(* IEC 61131-3 sources: 2026_Projet_YGO_ExcavatriceDragage/CODE_BACKUP/CODE_20260907_ChantierWeekEnd_v0.6.43/E_CODEURS, 7 files *)

(* ---- FB_Encoder.st ---- *)
(* =======================================================================
   🔌 FB_Encoder — Objet codeur complet (1 par treuil M1/M2)
   ───────────────────────────────────────────────────────────────
   🎯 Rôle : Regrouper toute la chaine codeur derriere une interface unique :
      Abs → Homing → Scale → Safety → Reliability → Speed.
   🔌 Frontiere hardware separee HwIn/HwOut (testable).
   🔒 Homing : autorise par HomingPermit (calcule par le caller), declenche
      par HomingAtTargetM (front). La cible est fournie par le caller.
   🔒 Fiabilite : gate EncoderFault (sans Homed) calcule AVANT Speed — purge
      de vitesse au meme scan. HomedAndReliable = gate strict interlock M3.
   🧩 Defaut : Fault:ST_Fault rempli par FB_FaultCore (instFault) depuis une liste
      de causes en clair (instCauses) — pattern FB_Joystick. Ready = Enable ET pas de
      defaut late. Interlocks machine sur les faits bruts, jamais sur Fault.Latched.
   📄 Doc : DOC/AF/AF_Partie-09_Fonction_Encoder_v2.4.md
   ======================================================================= *)

FUNCTION_BLOCK PUBLIC FB_Encoder
VAR_INPUT
    // === COMMANDES & AUTORISATIONS ===
    Enable                : BOOL;        // --> [CMD] Autorisation generale FB (TRUE=Autorise)
    Reset                 : BOOL;        // --> [CMD] Acquittement defaut (front montant)

    // === AUTORISATION HOMING (calculee par le caller PRG) ===
    HomingPermit          : BOOL;        // --> [CMD] TRUE = l'operateur a le droit de homer

    // === CONSIGNES HOMING ===
    HomingAtTargetM       : BOOL;        // --> [CMD] Demande homing vers cible (front montant)
    HomingAtZero          : BOOL;        // --> [CMD] Force homing a 0.0
    ConfirmCoherence      : BOOL;        // --> [CMD] Lever le doute d'incoherence boot
    CfgHomingTargetM      : REAL;        // --> [CFG] Cible libre homing unitaire (m)
    CfgTopSensorPosM      : REAL;        // --> [CFG] Cible homing nominal capteur haut (m)
    UseDynamicTarget      : BOOL;        // --> [CMD] Active cible dynamique
    DynamicHomingTargetM  : REAL;       // --> [CFG] Cible dynamique de referencement (m)

    // === CAPTEURS PHYSIQUES ===
    TopPositionSensor     : BOOL;        // --> [HW]  Capteur physique position haute unique

    // === BUS ETHERCAT & CAPTEUR HW (frontiere testable) ===
    HwIn                  : ST_fbEncoder_HwIn; // --> [HW] Retours hardware codeur

    // === MECANIQUE (constantes) ===
    PointsPerRev          : UDINT := 8192; // --> [CFG] Resolution codeur (pts/tour)
    CableM_PerRev         : REAL := 2.0;   // --> [CFG] Developpement cable par tour (m/tour)

    // === REGLAGES & CONFIGURATION ===
    Cfg                   : ST_fbEncoder_Cfg; // --> [CFG] Mode de confirmation preset
    PositionMinM          : REAL := -99.0; // --> [CFG] Plafond bornage physique bas (m)
    PositionMaxM          : REAL := 99.0;  // --> [CFG] Plafond bornage physique haut (m)
    BypassGlobal          : BOOL := FALSE; // --> [TST] Neutralisation defauts pour mise en service
END_VAR
VAR_OUTPUT
    // === ETATS IEC & SYNOPTIQUE ===
    Ready                 : BOOL;        // <-- [STAT] FB pret a fonctionner (Enable ET pas de defaut late)
    Fault                 : ST_Fault;    // <-- [DIAG] Brique defaut socle (live + latchee), remplie par FB_FaultCore

    // === FRONTIERE HW SORTIE (testable) ===
    HwOut                 : ST_fbEncoder_HwOut; // <-- [ACT] Ordres hardware codeur (preset)

    // === MESURES CONDITIONNEES (struct frontiere) ===
    Measurement           : ST_fbEncoder_Measurement; // <-- [BUS] Mesures + statuts (interface)

    // === ETATS CODEUR ===
    Homed                 : BOOL;        // <-- [STAT] Codeur reference (sortie homing)
    HomingSuspect         : BOOL;        // <-- [DIAG] Incoherence redemarrage a lever
    EncoderFault          : BOOL;        // <-- [SAFE] Gate general fiabilite (sans Homed)
    HomedAndReliable      : BOOL;        // <-- [STAT] Gate strict M3 : dispo ET ref ET pas incoherent
    PresetConfirmationFailed : BOOL;     // <-- [DIAG] Latch derniere verification preset echouee
END_VAR
VAR
    // === SOUS-INSTANCES FB (chaine codeur complete) ===
    instAbs        : FB_Encoder_Abs;          // * [INST] Acquisition brute codeur EtherCAT
    instHoming     : FB_Encoder_Homing;       // * [INST] Referencement (homing) nominal/unitaire
    instScale      : FB_Encoder_Scale;        // * [INST] Mise a l'echelle points -> metres
    instSafety     : FB_Encoder_Safety;       // * [INST] Bornage & coherence mesure
    instRel        : FB_EncoderReliability;   // * [INST] Gates de fiabilite
    instSpeed      : FB_Encoder_SpeedMeasure; // * [INST] Calcul vitesse cable
    instFault      : FB_FaultCore;            // * [INST] Socle de defaut (liste de causes -> ST_Fault)
    instCauses     : ARRAY[0..15] OF ST_FaultCause; // . [LOC] Liste des causes pour le socle FB_FaultCore
END_VAR
VAR_IN_OUT
    // === CALIBRATION PERSISTANTE (externe RETAIN, jamais membre) ===
    Calib                  : ST_Encoder_Calib; // <-> [BUS] Calibration RETAIN du treuil
END_VAR

{region "§1 Gate neutralisation"}
IF NOT Enable THEN
    Ready := FALSE;
    Measurement.RawPos := 0; Measurement.EncoderAvailable := FALSE;
    Measurement.CablePosM := 0.0; Measurement.CablePosMSafe := 0.0; Measurement.EncoderIncoherent := FALSE;
    Measurement.Speed_Mps := 0.0; Measurement.SignedSpeed_Mps := 0.0; Measurement.SpeedValid := FALSE;
    Measurement.HomingFault.Error := FALSE; Measurement.HomingFault.ErrorId := 0;
    Measurement.HomingLifecycle.Busy := FALSE; Measurement.HomingLifecycle.Done := FALSE;
    Measurement.AbsFault.Error := FALSE;    Measurement.AbsFault.ErrorId := 0;
    EncoderFault := TRUE;
    HomedAndReliable := FALSE;
    // Frontiere HW sortie : aucun ordre preset publie hors autorisation
    // (sinon PRG_02_Acquisition relaie une valeur perimee au codeur absolu -> preset parasite, reference corrompue)
    HwOut.PresetTriggerCmd := 0; HwOut.CodeSeqTriggerCmd := 0; HwOut.PresetValueOut := 0;
    // Reference connue MAINTENUE depuis Calib (RETAIN) meme FB desactive (AF09 §4) :
    // un FB desactive ne doit pas faire perdre la reference aux consommateurs aval (PRG_04, FB_Encoder_Scale).
    Homed := Calib.Homed;
    HomingSuspect := Calib.HomingSuspect;
    Measurement.HomingRefRaw := Calib.HomingRefRaw;
    // PresetConfirmationFailed est un diagnostic latch : il reste gele hors Enable
    // et ne doit pas etre efface par ce gate (AC3).
    // Socle appele meme Enable=FALSE : maintient le latch non acquitte et traite le Reset
    // hors autorisation (AC4). Les causes ne sont pas evaluees (Enable=FALSE -> vue live a 0),
    // les latches sont preserves.
    instFault(Enable := FALSE, Reset := Reset, Causes := instCauses);
    Fault := instFault.Fault;
    RETURN;
END_IF;
Ready := TRUE;
{endregion}

{region "§2 Abs"}
    instAbs(
    Enable              := Enable,
    Reset               := Reset,
    RawPosIn            := HwIn.RawPosIn,
    AlarmsIn            := HwIn.AlarmsIn,
    WarningsIn          := HwIn.WarningsIn,
    SlaveOperational    := HwIn.SlaveOperational,
    PresetRequest       := instHoming.PresetRequest,
    PresetValue         := instHoming.PresetValue,
    PointsPerRev        := PointsPerRev
);
{endregion}

{region "§3 Homing"}
instHoming(
    Enable               := Enable,
    Reset                := Reset,
    Home                 := HomingAtTargetM,
    HomingPermit         := HomingPermit,
    BtnConfirmCoherence  := ConfirmCoherence,
    UseDynamicTarget     := UseDynamicTarget,
    DynamicHomingTargetM := DynamicHomingTargetM,
    CfgHomingTargetM     := CfgHomingTargetM,
    CfgTopSensorPosM     := SEL(HomingAtZero, CfgTopSensorPosM, 0.0),
    TopPositionSensor    := TopPositionSensor,
    RawPos               := instAbs.RawPos,
    EncoderAvailable     := instAbs.EncoderAvailable,
    PresetStatusBit      := HwIn.PresetStatusBit,
    Cfg                  := Cfg,
    PointsPerRev         := PointsPerRev,
    MultiTurnRevsMax     := 4096,
    CableM_PerRev        := CableM_PerRev,
    BypassGlobal         := BypassGlobal,
    Calib                := Calib
);
{endregion}

{region "§4 Scale"}
instScale(
    RawPos       := instAbs.RawPos,
    HomingRefRaw := instHoming.HomingRefRaw,
    CableM_PerRev := CableM_PerRev,
    PointsPerRev := PointsPerRev
);
{endregion}

{region "§5 Safety"}
instSafety(
    Enable             := Enable,
    Reset              := Reset,
    CablePosM          := instScale.CablePosM,
    HomingSuspect      := instHoming.HomingSuspect,
    PositionMinM       := PositionMinM,
    PositionMaxM       := PositionMaxM,
    BypassGlobal       := BypassGlobal
);
{endregion}

{region "§6 Reliability"}
instRel(
    EncoderAvailable  := instAbs.EncoderAvailable,
    Homed             := instHoming.Homed,
    EncoderIncoherent := instSafety.EncoderIncoherent
);
{endregion}

{region "§7 Speed"}
instSpeed(
    Enable        := Enable,
    Reset         := Reset,
    SpdValueIn    := HwIn.SpdValueIn,
    PositionValid := NOT instRel.EncoderFault,
    CableM_PerRev := CableM_PerRev
);
{endregion}

{region "§8 Remplissage struct et synthese"}
Measurement.RawPos            := instAbs.RawPos;
Measurement.EncoderAvailable  := instAbs.EncoderAvailable;
Measurement.CablePosM         := instSafety.CablePosMSafe;
Measurement.CablePosMSafe     := instSafety.CablePosMSafe;
Measurement.EncoderIncoherent := instSafety.EncoderIncoherent;
Measurement.Speed_Mps         := instSpeed.Speed_Mps;
Measurement.SignedSpeed_Mps   := instSpeed.SignedSpeed_Mps;
Measurement.SpeedValid        := instSpeed.Valid;
Measurement.HomingFault        := instHoming.Fault;
Measurement.HomingLifecycle    := instHoming.Lifecycle;
Measurement.AbsFault           := instAbs.Fault;
Measurement.HomingRefRaw      := instHoming.HomingRefRaw;

// Frontiere HW sortie (preset)
HwOut.PresetTriggerCmd := instAbs.PresetTriggerCmd;
HwOut.CodeSeqTriggerCmd := instAbs.CodeSeqTriggerCmd;
HwOut.PresetValueOut    := instAbs.PresetValueOut;

// Etats codeur
Homed            := instHoming.Homed;
HomingSuspect    := instHoming.HomingSuspect;
EncoderFault     := instRel.EncoderFault;
HomedAndReliable := instRel.HomedAndReliable;
PresetConfirmationFailed := instHoming.PresetConfirmationFailed;

// Synthese statut facade : brique defaut socle (Fault:ST_Fault), pattern FB_Joystick.
// Causes exprimees en CLAIR (ST_FaultCause), alimentees UNIQUEMENT depuis les sorties
// publiques des sous-FB (encapsulation stricte, jamais de lecture VAR interne).
//   - Cause 0/1 : LIVE (Latching=FALSE) -> Fault.Error, retombe seule.
//   - Cause 2   : LATCHED (Latching=TRUE) -> arme Fault.Latched, acquittee au Reset front.
// Interlock machine toujours sur les faits bruts (EncoderFault, HomedAndReliable,
// EncoderIncoherent), jamais sur Fault.Latched (conservation).
instCauses[0].Active := NOT instAbs.EncoderAvailable; instCauses[0].Latching := FALSE;
instCauses[0].Texte := 'Perte materiel / communication codeur EtherCAT';
instCauses[1].Active := instSafety.EncoderIncoherent; instCauses[1].Latching := FALSE;
instCauses[1].Texte := 'Incoherence mesure / saut de position codeur';
instCauses[2].Active := instHoming.PresetConfirmationFailed; instCauses[2].Latching := TRUE;
instCauses[2].Texte := 'Echec confirmation transaction preset codeur';

// Socle appele APRES le pipeline : causes du scan courant, aucun scan de retard (AC4).
instFault(Enable := Enable, Reset := Reset, Causes := instCauses);
Fault := instFault.Fault;     // source de verite = socle
Ready := Enable AND NOT Fault.Latched;
{endregion}

(* ---- FB_Encoder_Abs.st ---- *)
(* =======================================================================
   🔌 FB_Encoder_Abs — Acquisition codeur absolu (accès bus EtherCAT)
   ───────────────────────────────────────────────────────────────
   🎯 Rôle : Accès bus EtherCAT, extraction positions brutes et séquence de Preset SDO
   🔒 Polarité : EncoderAvailable=TRUE si communication bus et esclave OK
   🔌 Architecture : Module d'acquisition codeur absolu
   📄 Doc métier : DOC/AF/AF_Partie-09_Fonction_Encoder_v2.4.md
   ======================================================================= *)

// === DECLARATION (à coller dans la partie déclaration du POU FB_Encoder_Abs) ===

FUNCTION_BLOCK PUBLIC FB_Encoder_Abs
VAR_INPUT
    // === COMMANDES & AUTORISATIONS ===
    Enable              : BOOL;        // --> [CMD] Autorisation generale FB (TRUE=Autorise)
    Reset               : BOOL;        // --> [CMD] Acquittement defaut (front montant)
    PresetRequest       : BOOL;        // --> [CMD] Demande de preset (front montant)

    // === BUS ETHERCAT & CAPTEUR HW ===
    RawPosIn            : UDINT;       // --> [HW]  Position brute EtherCAT
    AlarmsIn            : UINT;        // --> [HW]  Codes alarmes bruts EtherCAT
    WarningsIn          : UINT;        // --> [HW]  Codes avertissements bruts EtherCAT
    SlaveOperational    : BOOL;        // --> [HW]  Statut esclave EtherCAT operationnel

    // === PARAMETRES & REGLAGES ===
    PointsPerRev        : UDINT := 8192; // --> [CFG] Resolution codeur (pts/tour)
    PresetValue         : UDINT;       // --> [CFG] Valeur cible de preset
    PresetTimeout       : TIME := T#2s;// --> [CFG] Temporisation max attente preset
    PresetTolerancePts  : UDINT := 10; // --> [CFG] Tolerance relecture post-preset (pts)
END_VAR
VAR_OUTPUT
    // === ETATS IEC & SYNOPTIQUE ===
    Ready               : BOOL;        // <-- [STAT] FB pret a fonctionner
    // 🧩 Statut transverse (forme cible ST_Fault)
    Fault               : ST_Fault;

    // === MESURES & DONNEES CODEUR ===
    RawPos              : UDINT;       // <-- [DIAG] Position brute gelee si non disponible
    EncoderAvailable    : BOOL;        // <-- [STAT] Codeur operationnel et disponible
    AngleRaw            : UINT;        // <-- [DIAG] Angle brut sur un tour (MOD PointsPerRev)
    TurnCount           : UDINT;       // <-- [DIAG] Nombre de tours bruts (RawPos / PointsPerRev)

    // === COMMANDES & ECHANGE BUS ETHERCAT ===
    PresetTriggerCmd    : WORD;        // <-- [ACT]  Ordre declenchement preset vers PDO Rx
    CodeSeqTriggerCmd   : WORD;        // <-- [ACT]  Ordre sequence code vers PDO Rx
    PresetValueOut      : UDINT;       // <-- [ACT]  Valeur de preset transmise au PDO Rx
END_VAR
VAR
    // === DETECTEURS DE FRONT ===
    ResetEdge           : R_TRIG;      // . [LOC] Detecteur front montant Reset
    PresetReqEdge       : R_TRIG;      // . [LOC] Detecteur front montant PresetRequest

    // === TEMPORISATEURS INTERNES ===
    PresetTimer         : TON;         // . [LOC] Temporisateur timeout sequence preset
    PresetTimerVisual   : TON;         // . [LOC] Temporisateur maintien visuel impulsion (500ms)

    // === VARIABLES INTERNES DE CALCUL & ETAT ===
    PresetSeqStep       : INT;         // . [LOC] Etape sequence preset (0:IDLE, 1:PULSE/WAIT)
    RawDiff             : DINT;        // . [LOC] Ecart signe entre RawPos et PresetValueOut
    PresetCompleted     : BOOL;        // . [LOC] Fait de fin de maintien preset (un scan)
    PresetTimeoutError  : BOOL;        // . [LOC] Latch interne timeout séquence preset

    // === SOCLE DEFAUT (FB_FaultCore) ===
    instFault           : FB_FaultCore;                   // * [INST] Socle défaut transverse
    instCauses          : ARRAY[0..15] OF ST_FaultCause;  // . [LOC] Table des causes nommées
END_VAR

// === IMPLEMENTATION (à coller dans le corps ST du POU FB_Encoder_Abs) ===

{region "§1 Causes & Socle Défaut (évalué en continu)"}
// 🔑 1. RESET FRONT
ResetEdge(CLK := Reset);

// 🔍 2. DIAGNOSTIC BUS / ALARME (Cause 0 : live)
instCauses[0].Active   := (AlarmsIn <> 0) OR NOT SlaveOperational;
instCauses[0].Latching := FALSE;
instCauses[0].Texte    := 'Defaut communication EtherCAT codeur absolu';

// ⏱️ 3. TIMEOUT PRESET (Cause 1 : latched)
IF ResetEdge.Q AND (PresetSeqStep = 0) THEN
    PresetTimeoutError := FALSE;
END_IF;
instCauses[1].Active   := PresetTimeoutError;
instCauses[1].Latching := TRUE;
instCauses[1].Texte    := 'Timeout sequence preset SDO codeur';

// Appel du socle de défaut
instFault(Enable := Enable, Reset := Reset, Causes := instCauses);
Fault := instFault.Fault;

EncoderAvailable := NOT instCauses[0].Active;
{endregion}

{region "§2 Gate neutralisation"}
// 🛑 2. GATE
IF NOT Enable THEN
    EncoderAvailable := FALSE;
    Ready := FALSE;
    PresetTriggerCmd := 0; CodeSeqTriggerCmd := 0; PresetValueOut := 0;
    PresetSeqStep := 0;
    PresetCompleted := FALSE;
    PresetTimer(IN := FALSE, PT := PresetTimeout);
    PresetTimerVisual(IN := FALSE, PT := T#500MS);
    // RawPos, AngleRaw et TurnCount sont volontairement gelés hors Enable
    // (AF09 F09.01 / AC5) : aucune lecture bus ni remise a zero dans ce gate.
    RETURN;
END_IF;

Ready := Enable AND NOT Fault.Latched;
{endregion}

{region "§3 Lecture position"}
// 📥 3. LECTURE POSITION — GELER SUR DOUTE (Partie10 §6)
// Si EncoderAvailable=FALSE : RawPos/AngleRaw/TurnCount conservent leur dernière valeur (pas de RETURN
// global ici pour ne pas geler aussi la séquence preset/l'état — seule la lecture est gelée).
IF EncoderAvailable THEN
    RawPos := RawPosIn;   // Sens de comptage géré côté codeur (CoE 6000h bit0, startup parameter CODESYS) — voir Partie10 §3bis. Plus de calcul ici.
    AngleRaw := UDINT_TO_UINT(RawPos MOD PointsPerRev);
    TurnCount := RawPos / PointsPerRev;
END_IF;
{endregion}

{region "§4 Séquence preset"}
// 🔧 4. SÉQUENCE PRESET (écriture bus)
// PresetTriggerCmd := 2 déclenche le référencement à PresetValue (valeur de commande, pas un
// masque de bits). CodeSeqTriggerCmd : rôle non identifié — laissé à 0, PAS piloté tant que sa
// fonction n'est pas confirmée. Ne jamais lui donner une valeur arbitraire.
PresetReqEdge(CLK := PresetRequest);
PresetCompleted := FALSE;
CodeSeqTriggerCmd := 0;                 // non piloté — rôle inconnu, voir note ci-dessus
CASE PresetSeqStep OF
    0: // IDLE
        PresetTriggerCmd := 0;
        IF PresetReqEdge.Q AND EncoderAvailable THEN
            PresetValueOut := PresetValue;
            PresetSeqStep := 1;
            PresetTimer(IN := TRUE, PT := PresetTimeout);
        END_IF;
    1: // Déclenchement preset (laissé actif pendant 0.5s pour confort visuel en simulation/bus)
        PresetTriggerCmd := 2;   // Référence le codeur à PresetValueOut
        RawDiff := UDINT_TO_DINT(RawPos) - UDINT_TO_DINT(PresetValueOut);
        IF ABS(RawDiff) <= UDINT_TO_DINT(PresetTolerancePts) THEN
            PresetTimer(IN := FALSE, PT := PresetTimeout);
            PresetTimerVisual(IN := TRUE, PT := T#500MS);
            IF PresetTimerVisual.Q THEN
                PresetTriggerCmd := 0;
                PresetCompleted := TRUE;
                PresetSeqStep := 0;
                PresetTimerVisual(IN := FALSE, PT := T#500MS);
            END_IF;
        ELSIF PresetTimer.Q THEN
            PresetTriggerCmd := 0;
            PresetTimeoutError := TRUE;
            PresetSeqStep := 0;
            PresetTimer(IN := FALSE, PT := PresetTimeout);
            PresetTimerVisual(IN := FALSE, PT := T#500MS);
        END_IF;
END_CASE;
{endregion}

(* ---- FB_Encoder_Homing.st ---- *)
(* =======================================================================
   ⚙️ FB_Encoder_Homing — Référencement codeur nominal ou unitaire
   ───────────────────────────────────────────────────────────────
   🎯 Rôle : Séquence de référencement nominal (capteur haut) ou unitaire (MAINT_N2)
   🔒 Polarité : Homed=TRUE dès qu'un référencement valide est enregistré
   🔌 Architecture : Expose ST_Encoder_Calib en VAR_IN_OUT
   📄 Doc métier : DOC/AF/AF_Partie-09_Fonction_Encoder_v2.4.md
   ======================================================================= *)

// === DECLARATION (à coller dans la partie déclaration du POU FB_Encoder_Homing) ===

FUNCTION_BLOCK PUBLIC FB_Encoder_Homing
VAR_INPUT
    // === COMMANDES & AUTORISATIONS ===
    Enable                 : BOOL;        // --> [CMD] Autorisation generale FB (TRUE=Autorise)
    Reset                  : BOOL;        // --> [CMD] Acquittement defaut (front montant)
    Home                   : BOOL;        // --> [CMD] Demande de referencement (front)
    HomingPermit           : BOOL;        // --> [CMD] Autorisation de homer (calculee par le caller)
    BtnConfirmCoherence    : BOOL;        // --> [CMD] Levee de doute d'incoherence au boot (front)

    // === CIBLES & CONFIGURATION HOMING ===
    CfgHomingTargetM       : REAL;        // --> [CFG] Cible libre homing unitaire (m)
    UseDynamicTarget       : BOOL := FALSE; // --> [CFG] Activation cible dynamique
    DynamicHomingTargetM   : REAL := 0.0; // --> [CFG] Cible dynamique de referencement (m)
    CfgTopSensorPosM       : REAL := 8.5; // --> [CFG] Cible homing nominal capteur haut (m)

    // === RETOURS HW & CAPTEURS ===
    TopPositionSensor      : BOOL;        // --> [HW]  Capteur physique position haute unique
    // === MESURES & RETOURS FB CODEUR ABSOLU ===
    RawPos                 : UDINT;       // --> [HW]  Position brute codeur (sortie FB_Encoder_Abs)
    EncoderAvailable       : BOOL;        // --> [HW]  Codeur absolu disponible et valide
    PresetStatusBit        : BOOL;        // --> [HW]  Bit d'etat preset optionnel, FALSE si non cable

    // === REGLAGES TRANSACTION PRESET ===
    Cfg                    : ST_fbEncoder_Cfg; // --> [CFG] Mode de confirmation preset

    // === CARACTERISTIQUES MECANIQUES & BUS ===
    PointsPerRev           : UDINT := 8192; // --> [CFG] Resolution codeur (pts/tour)
    MultiTurnRevsMax       : UDINT := 4096; // --> [CFG] Capacite multitour max codeur (tours)
    CableM_PerRev          : REAL := 2.0;   // --> [CFG] Perimetre tambour / developpement cable (m/tour)

    // === TESTS & BYPASS ===
    BypassGlobal           : BOOL := FALSE; // --> [TST] Neutralisation securites pour mise en service
END_VAR
VAR_OUTPUT
    // === ETATS IEC & SYNOPTIQUE ===
    Ready                  : BOOL;        // <-- [STAT] FB pret a fonctionner
    // 🧩 Statut transverse (forme cible ST_Fault)
    Fault                  : ST_Fault;
    // 🧩 Cycle de vie (forme cible ST_Lifecycle)
    Lifecycle              : ST_Lifecycle;

    // === COMMANDES VERS FB_ENCODER_ABS ===
    PresetRequest          : BOOL;        // <-- [ACT]  Pulse demande d'ecriture preset SDO
    PresetValue            : UDINT;       // <-- [ACT]  Valeur de cible brute pour preset SDO

    // === RESULTATS & MEMOIRE CALIBRATION ===
    Homed                  : BOOL;        // <-- [STAT] Codeur pagine et referencie
    HomingSuspect          : BOOL;        // <-- [DIAG] Incoherence redemarrage a lever
    HomingRefRaw           : UDINT;       // <-- [DIAG] Offset de reference brut calcule
    PresetConfirmationFailed : BOOL;      // <-- [DIAG] Latch derniere verification preset echouee
END_VAR
VAR_IN_OUT
    // === STRUCTURE DE CALIBRATION PERSISTANTE ===
    Calib                  : ST_Encoder_Calib; // <-> [BUS] Structure de calibration RETAIN
END_VAR
VAR
    // === DETECTEURS DE FRONT ===
    ResetEdge              : R_TRIG;      // . [LOC] Detecteur front montant Reset
    HomeEdge               : R_TRIG;      // . [LOC] Detecteur front montant Home
    ConfirmCoherenceEdge   : R_TRIG;      // . [LOC] Detecteur front montant BtnConfirmCoherence
    TopSensorEdge          : R_TRIG;      // . [LOC] Detecteur front montant TopPositionSensor
    DynamicTargetEdge      : R_TRIG;      // . [LOC] Detecteur front montant UseDynamicTarget

    // === ETATS & DRAPEAUX INTERNES ===
    InitDone               : BOOL;        // . [LOC] Controle incoherence boot effectue
    HomingModeOk           : BOOL;        // . [LOC] Mode de fonctionnement valide pour homing
    NominalHomingTrigger   : BOOL;        // . [LOC] Condition de declenchement homing nominal
    UnitaryHomingTrigger   : BOOL;        // . [LOC] Condition de declenchement homing unitaire
    DynamicHomingTrigger   : BOOL;        // . [LOC] Condition de declenchement homing dynamique
    HomingTrigger          : BOOL;        // . [LOC] Synthese declenchement homing
    PresetVerificationActive : BOOL;      // . [LOC] Verification preset en attente
    PresetConfirmed        : BOOL;        // . [LOC] Resultat du mode de confirmation selectionne

    // === DRAPEAUX DEFAUTS INTERNES ===
    HomingModeError        : BOOL;        // . [LOC] Latch erreur mode
    TargetOutOfRangeError  : BOOL;        // . [LOC] Latch cible hors limites
    PresetFailError        : BOOL;        // . [LOC] Latch échec preset
    BootIncoherentError    : BOOL;        // . [LOC] Latch incohérence boot

    // === VARIABLES DE CALCUL ===
    TargetPoints           : DINT;        // . [LOC] Ecart cible converti en points
    TargetPositionM        : REAL;        // . [LOC] Cible retenue en metres
    RawDiffRestart         : DINT;        // . [LOC] Ecart brut de position au redemarrage
    PendingHomingRefRaw    : UDINT;       // . [LOC] Reference candidate, non publiee avant succes
    CandidateRawDiff       : DINT;        // . [LOC] Ecart brut de la mesure candidate
    CandidateCablePosM     : REAL;        // . [LOC] Position candidate calculee avant commit
    ReadbackOk             : BOOL;        // . [LOC] Mesure candidate dans la tolerance
    StatusBitOk            : BOOL;        // . [LOC] Etat du bit optionnel de confirmation
    PresetVerifyTimer      : TON;         // . [LOC] Temporisation historique de verification 500ms

    // === SOCLE DEFAUT (FB_FaultCore) ===
    instFault              : FB_FaultCore;                   // * [INST] Socle défaut transverse
    instCauses             : ARRAY[0..15] OF ST_FaultCause;  // . [LOC] Table des causes nommées
END_VAR

VAR CONSTANT
    // === TOLERANCE & TEMPORISATION TRANSACTION ===
    CST_HomingVerifyToleranceM : REAL := 0.010; // Tolerance mesure cible (m)
    CST_PresetVerifyTime        : TIME := T#50MS; // Latence historique avant relecture
END_VAR

// === IMPLEMENTATION (à coller dans le corps ST du POU FB_Encoder_Homing) ===

{region "§1 Causes & Socle Défaut (évalué en continu)"}
// 🔑 1. FRONTS
ResetEdge(CLK := Reset);
HomeEdge(CLK := Home);
ConfirmCoherenceEdge(CLK := BtnConfirmCoherence);

// Effacement des latches d'erreur sur Reset conscient
IF ResetEdge.Q THEN
    PresetConfirmationFailed := FALSE;
    HomingModeError := FALSE;
    TargetOutOfRangeError := FALSE;
    PresetFailError := FALSE;
END_IF;

// Levée de doute incohérence boot (BtnConfirmCoherence)
IF ConfirmCoherenceEdge.Q AND HomingPermit THEN
    Calib.HomingSuspect := FALSE;
    BootIncoherentError := FALSE;
END_IF;

// Configuration des causes nommées
instCauses[0].Active   := HomingModeError;
instCauses[0].Latching := TRUE;
instCauses[0].Texte    := 'Homing non autorise dans ce mode';

instCauses[1].Active   := TargetOutOfRangeError;
instCauses[1].Latching := TRUE;
instCauses[1].Texte    := 'Cible de homing hors plage';

instCauses[2].Active   := PresetFailError;
instCauses[2].Latching := TRUE;
instCauses[2].Texte    := 'Echec confirmation transaction preset';

instCauses[3].Active   := BootIncoherentError;
instCauses[3].Latching := TRUE;
instCauses[3].Texte    := 'Incoherence position codeur au demarrage';

// Appel du socle de défaut
instFault(Enable := Enable, Reset := Reset, Causes := instCauses);
Fault := instFault.Fault;
{endregion}

{region "§2 Gate neutralisation"}
// 🛑 2. GATE — neutralisation ; on continue toutefois d'exposer le dernier état RETAIN connu
// (FB_Encoder_Scale a besoin de HomingRefRaw même si ce FB est désactivé)
IF NOT Enable THEN
    PresetRequest := FALSE;
    PresetValue := 0;
    Ready := FALSE;
    Lifecycle.Busy := FALSE;
    Lifecycle.Done := FALSE;
    InitDone := FALSE;   // Force un nouveau contrôle à la prochaine activation
    PresetVerificationActive := FALSE;
    PresetVerifyTimer(IN := FALSE, PT := CST_PresetVerifyTime);
    Homed := Calib.Homed;
    HomingSuspect := Calib.HomingSuspect;
    HomingRefRaw := Calib.HomingRefRaw;
    // PresetConfirmationFailed est un diagnostic latch : il est gelé hors Enable
    RETURN;
END_IF;

Ready := Enable AND NOT Fault.Latched;
{endregion}

{region "§3 Cohérence au redémarrage"}
// 🔍 3. COHÉRENCE AU REDÉMARRAGE — une fois par session Enable, dès que le codeur répond
IF NOT InitDone THEN
    IF EncoderAvailable THEN
        RawDiffRestart := UDINT_TO_DINT(RawPos) - UDINT_TO_DINT(Calib.LastKnownRawPos);
        IF Calib.Homed AND (ABS(RawDiffRestart) > UDINT_TO_DINT(Calib.RestartCoherenceTolerancePts)) THEN
            Calib.HomingSuspect := TRUE;
            BootIncoherentError := TRUE;
        END_IF;
        InitDone := TRUE;
    END_IF;
END_IF;
{endregion}

{region "§4 Demande et déclenchement homing"}
// ⚙️ 4. DEMANDE & DÉCLENCHEMENT HOMING
PresetRequest := FALSE;
PresetValue := 0;
TopSensorEdge(CLK := TopPositionSensor);
DynamicTargetEdge(CLK := UseDynamicTarget);

HomingModeOk := HomingPermit;

IF HomeEdge.Q AND NOT HomingModeOk THEN
    HomingModeError := TRUE;
END_IF;

NominalHomingTrigger := HomingModeOk AND NOT UseDynamicTarget
                         AND ((Home AND TopSensorEdge.Q) OR (HomeEdge.Q AND TopPositionSensor));

UnitaryHomingTrigger := HomingModeOk AND NOT UseDynamicTarget AND HomeEdge.Q;

DynamicHomingTrigger := HomingModeOk AND (DynamicTargetEdge.Q OR (UseDynamicTarget AND HomeEdge.Q));

HomingTrigger := (NominalHomingTrigger OR UnitaryHomingTrigger OR DynamicHomingTrigger)
                 AND NOT PresetVerificationActive;

IF HomingTrigger THEN
    IF UseDynamicTarget THEN
        TargetPositionM := DynamicHomingTargetM;
    ELSIF NominalHomingTrigger THEN
        TargetPositionM := CfgTopSensorPosM;
    ELSE
        TargetPositionM := CfgHomingTargetM;
    END_IF;

    // Bornage obligatoire avant écriture (CODE_QUALITY_STANDARDS §6) [-99;+99] m
    IF (TargetPositionM < -99.0) OR (TargetPositionM > 99.0) THEN
        TargetOutOfRangeError := TRUE;
    ELSE
        TargetPoints := REAL_TO_DINT(TargetPositionM * UDINT_TO_REAL(PointsPerRev) / CableM_PerRev);
        PendingHomingRefRaw := DINT_TO_UDINT(UDINT_TO_DINT(RawPos) - TargetPoints);
        PresetValue := RawPos;
        PresetRequest := TRUE;
        PresetVerificationActive := TRUE;
        Lifecycle.Done := FALSE;
    END_IF;
END_IF;
{endregion}

{region "§5 Suivi de transaction preset"}
// ⏳ 5. SUIVI DE LA TRANSACTION PRESET
PresetVerifyTimer(IN := PresetVerificationActive, PT := CST_PresetVerifyTime);
IF PresetVerificationActive AND PresetVerifyTimer.Q THEN
    CandidateRawDiff := UDINT_TO_DINT(RawPos) - UDINT_TO_DINT(PendingHomingRefRaw);
    IF PointsPerRev <> 0 THEN
        CandidateCablePosM := DINT_TO_REAL(CandidateRawDiff) * CableM_PerRev / UDINT_TO_REAL(PointsPerRev);
    ELSE
        CandidateCablePosM := 0.0;
    END_IF;
    ReadbackOk := ABS(CandidateCablePosM - TargetPositionM) <= CST_HomingVerifyToleranceM;
    StatusBitOk := PresetStatusBit;

    CASE Cfg.PresetConfirmMode OF
        E_PresetConfirmMode.READBACK_ONLY:
            PresetConfirmed := ReadbackOk;
        E_PresetConfirmMode.READBACK_AND_STATUSBIT:
            PresetConfirmed := ReadbackOk AND StatusBitOk;
        E_PresetConfirmMode.STATUSBIT_ONLY:
            PresetConfirmed := StatusBitOk;
        ELSE
            PresetConfirmed := FALSE;
    END_CASE;

    IF PresetConfirmed THEN
        Calib.HomingRefRaw := PendingHomingRefRaw;
        Calib.Homed := TRUE;
        Calib.HomingSuspect := FALSE;
        Calib.LastKnownRawPos := RawPos;
        PresetConfirmationFailed := FALSE;
        PresetFailError := FALSE;
        Lifecycle.Done := TRUE;
    ELSE
        Calib.HomingSuspect := TRUE;
        PresetConfirmationFailed := TRUE;
        PresetFailError := TRUE;
        Lifecycle.Done := FALSE;
    END_IF;

    PresetVerificationActive := FALSE;
    PresetVerifyTimer(IN := FALSE, PT := CST_PresetVerifyTime);
END_IF;
{endregion}

{region "§6 Sorties état & calibration"}
// 📤 6. SORTIES ÉTAT & CALIBRATION
IF EncoderAvailable AND NOT PresetVerificationActive THEN
    Calib.LastKnownRawPos := RawPos;
END_IF;

Lifecycle.Busy := PresetVerificationActive;
Homed := Calib.Homed AND NOT Calib.HomingSuspect;
HomingSuspect := Calib.HomingSuspect;
HomingRefRaw := Calib.HomingRefRaw;
{endregion}

(* ---- FB_Encoder_Safety.st ---- *)
(* =======================================================================
   🛡️ FB_Encoder_Safety — Bornage physique & surveillance cohérence
   ───────────────────────────────────────────────────────────────
   🎯 Rôle : Bornage physique absolu [-99; +99]m et relais d'incohérence redémarrage
   🔒 Polarité : EncoderIncoherent=TRUE en cas de hors bornes ou HomingSuspect
   🛡️ Sécurité : Verrouillage de la position câble sûre
   📄 Doc métier : DOC/AF/AF_Partie-09_Fonction_Encoder_v2.4.md
   ======================================================================= *)

FUNCTION_BLOCK PUBLIC FB_Encoder_Safety
VAR_INPUT
    // === COMMANDES & AUTORISATIONS ===
    Enable                : BOOL;        // --> [CMD] Autorisation generale FB (TRUE=Autorise)
    Reset                 : BOOL;        // --> [CMD] Acquittement defaut (front montant)

    // === MESURES & ALERTE HOMING ===
    CablePosM             : REAL;        // --> [HW]  Position calculee (m, sortie FB_Encoder_Scale)
    HomingSuspect         : BOOL;        // --> [SAFE] Alerte incoherence redemarrage (FB_Encoder_Homing)

    // === REGLAGES & BORNES PHYSIQUES ===
    PositionMinM          : REAL := -99.0; // --> [CFG] Plafond bornage physique bas (m)
    PositionMaxM          : REAL := 99.0;  // --> [CFG] Plafond bornage physique haut (m)

    // === TESTS & BYPASS ===
    BypassGlobal          : BOOL := FALSE; // --> [TST] Neutralisation defaut de bornage pour mise en service
END_VAR
VAR_OUTPUT
    // === ETATS IEC & SYNOPTIQUE ===
    Ready                 : BOOL;        // <-- [STAT] FB pret a fonctionner
    // 🧩 Statut transverse (forme cible ST_Fault)
    Fault                 : ST_Fault;

    // === MESURES SURE & SECURITE ===
    CablePosMSafe         : REAL;        // <-- [DIAG] Position cable instantanee transmise (m)
    EncoderIncoherent     : BOOL;        // <-- [SAFE] Incoherence ou hors bornes (TRUE = defaut)
END_VAR
VAR
    // === DETECTEURS DE FRONT ===
    ResetEdge             : R_TRIG;      // . [LOC] Detecteur front montant Reset

    // === SOCLE DEFAUT (FB_FaultCore) ===
    instFault             : FB_FaultCore;                   // * [INST] Socle défaut transverse
    instCauses            : ARRAY[0..15] OF ST_FaultCause;  // . [LOC] Table des causes nommées
END_VAR

// === IMPLEMENTATION ===

{region "§1 Causes & Socle Défaut (évalué en continu)"}
// 🔑 1. RESET FRONT
ResetEdge(CLK := Reset);

// 🔍 2. SURVEILLANCE BORNAGE & INCOHÉRENCE BOOT
instCauses[0].Active   := NOT BypassGlobal AND ((CablePosM < PositionMinM) OR (CablePosM > PositionMaxM));
instCauses[0].Latching := FALSE;
instCauses[0].Texte    := 'Depassement bornes physiques absolues cable';

instCauses[1].Active   := NOT BypassGlobal AND HomingSuspect;
instCauses[1].Latching := FALSE;
instCauses[1].Texte    := 'Incoherence position au redemarrage';

// Appel du socle de défaut
instFault(Enable := Enable, Reset := Reset, Causes := instCauses);
Fault := instFault.Fault;
{endregion}

{region "§2 Gate neutralisation"}
// 🛑 2. GATE
IF NOT Enable THEN
    Ready := FALSE;
    CablePosMSafe := CablePosM;
    EncoderIncoherent := FALSE;
    RETURN;
END_IF;

Ready := Enable AND NOT Fault.Latched;
{endregion}

{region "§3 Transmission mesure et sécurité"}
// 📏 3. TRANSMISSION DE LA MESURE & SÉCURITÉ
CablePosMSafe := CablePosM;
EncoderIncoherent := Fault.Error;
{endregion}

(* ---- FB_Encoder_Scale.st ---- *)
(* =======================================================================
   ⚙️ FB_Encoder_Scale — Mise à l'échelle points → mètres (1 par treuil)
   ───────────────────────────────────────────────────────────────
   🎯 Rôle : Calcul de la position câble en mètres par conversion arithmétique signée
   🔒 Polarité : CablePosM signée (+ enroulé, - sous l'eau)
   🔌 Architecture : Convertisseur de mesure unitaire par treuil
   📄 Doc métier : DOC/AF/AF_Partie-09_Fonction_Encoder_v2.4.md
   ======================================================================= *)

// === DECLARATION (à coller dans la partie déclaration du POU FB_Encoder_Scale) ===

FUNCTION_BLOCK PUBLIC FB_Encoder_Scale
VAR_INPUT
    // === DONNEES ENTREE & REFERENCES BRUTES ===
    RawPos          : UDINT;       // --> [HW]  Position brute codeur (sortie FB_Encoder_Abs, gelee sur doute)
    HomingRefRaw    : UDINT;       // --> [CFG] Reference brute figee au dernier homing (ST_Encoder_Calib)

    // === PARAMETRES & RATIOS DE CONVERSION ===
    CableM_PerRev   : REAL := 2.0; // --> [CFG] Developpement cable par tour tambour (m/tour)
    PointsPerRev    : UDINT := 8192;// --> [CFG] Resolution codeur (pts/tour)
END_VAR
VAR_OUTPUT
    // === MESURE CONVERTIE ===
    CablePosM       : REAL;        // <-- [DIAG] Position cable en metres (+ enroule, - sous l'eau)
END_VAR
VAR
    // === CALCULS INTERNES ===
    RawDiff         : DINT;        // . [LOC] Ecart signe RawPos - HomingRefRaw
END_VAR

// === IMPLEMENTATION (à coller dans le corps ST du POU FB_Encoder_Scale) ===

// 🧮 Écart signé sûr : conversion DINT AVANT soustraction (§3.1) — jamais l'inverse
RawDiff := UDINT_TO_DINT(RawPos) - UDINT_TO_DINT(HomingRefRaw);

// 📏 Formule fixe points → mètres (Partie10 §2), garde division par zéro
IF PointsPerRev > 0 THEN
    CablePosM := DINT_TO_REAL(RawDiff) * (CableM_PerRev / UDINT_TO_REAL(PointsPerRev));
ELSE
    CablePosM := 0.0;
END_IF;

(* ---- FB_Encoder_SpeedMeasure.st ---- *)
(* =======================================================================
   ⚙️ FB_Encoder_SpeedMeasure — Mesure de vitesse câble directe codeur
   ───────────────────────────────────────────────────────────────
   🎯 Rôle : Conversion directe du mot de vitesse natif codeur EtherCAT (m/s)
   ⚙️ Source CoE : Objet 0x6031:01 en 0.1 RPM (dixième de tour/min)
   📐 Formule : V(m/s) = (SpdValue * 0.1 * CableM_PerRev) / 60.0
   🛡️ Sans bornage : zéro clamping artificiel, suppression délai filtre PT1
   📄 Doc métier : DOC/AF/AF_Partie-09_Fonction_Encoder_v2.4.md
   ======================================================================= *)

FUNCTION_BLOCK PUBLIC FB_Encoder_SpeedMeasure
VAR_INPUT
    // === COMMANDES & AUTORISATIONS ===
    Enable              : BOOL;        // --> [CMD] Autorisation generale FB (TRUE=Autorise)
    Reset               : BOOL;        // --> [CMD] Purge immediate (front montant)

    // === MESURES EN ENTREE ===
    SpdValueIn          : DINT;        // --> [HW]  Mot de vitesse brut EtherCAT (0x6031:01 en 0.1 RPM)
    PositionValid       : BOOL;        // --> [SAFE] Validite de la chaine codeur
    CableM_PerRev       : REAL := 2.0; // --> [CFG] Developpement cable par tour tambour (m/tour)
END_VAR
VAR_OUTPUT
    // === VITESSE CÂBLE QUALIFIÉE (m/s) ===
    Speed_Mps           : REAL;        // <-- [DIAG] Vitesse absolue directe (m/s)
    SignedSpeed_Mps     : REAL;        // <-- [DIAG] Vitesse signee directe (+ montee, - descente) (m/s)
    Valid               : BOOL;        // <-- [STAT] Validite mesure (TRUE si codeur operationnel et autorise)
END_VAR
VAR
    // === MEMOIRES & DETECTEURS ===
    ResetEdge           : R_TRIG;      // . [LOC] Detecteur front montant Reset
END_VAR

{region "§1 Gate de neutralisation & Reset"}
ResetEdge(CLK := Reset);

// Purge immediate sur perte de confiance, desactivation ou Reset
IF NOT Enable OR ResetEdge.Q OR NOT PositionValid THEN
    Speed_Mps       := 0.0;
    SignedSpeed_Mps := 0.0;
    Valid           := FALSE;
    RETURN;
END_IF;
{endregion}

{region "§2 Conversion directe vitesse CoE (0.1 RPM -> m/s)"}
// Formule cinematique directe :
// N_RPM = SpdValueIn * 0.1
// V_mps = (N_RPM * CableM_PerRev) / 60.0 = (DINT_TO_REAL(SpdValueIn) * 0.1 * CableM_PerRev) / 60.0
SignedSpeed_Mps := (DINT_TO_REAL(SpdValueIn) * 0.1 * CableM_PerRev) / 60.0;
Speed_Mps       := ABS(SignedSpeed_Mps);
Valid           := TRUE;
{endregion}

END_FUNCTION_BLOCK

(* ---- FB_EncoderReliability.st ---- *)
(* =======================================================================
   🛡️ FB_EncoderReliability — Gates de fiabilite de la chaine codeur
   ───────────────────────────────────────────────────────────────
   🎯 Rôle : Synthetise les gates de fiabilite d'un treuil a partir des
      faits produits par la chaine codeur (Abs/Homing/Safety), pur calcul
      combinatoire, sans memoire ni machine d'etat.
   🔒 Polarité :
      EncoderFault     = NOT EncoderAvailable OR EncoderIncoherent   (gate GENERAL, SANS Homed)
      HomedAndReliable = EncoderAvailable AND Homed AND NOT EncoderIncoherent (gate STRICT M3)
   🧩 Responsabilite scindee (D-A2bis) : Homing = referencement, Safety = coherence,
      ce FB = « le codeur est fiable ». Aucune recomposition chez les consommateurs.
   📄 Doc : DOC/AF/AF_Partie-09_Fonction_Encoder_v2.4.md
   ======================================================================= *)

FUNCTION_BLOCK PUBLIC FB_EncoderReliability
VAR_INPUT
    // === FAITS DE LA CHAINE CODEUR ===
    EncoderAvailable  : BOOL;        // --> [HW]  Codeur operationnel sur bus (FB_Encoder_Abs)
    Homed             : BOOL;        // --> [STAT] Codeur reference (FB_Encoder_Homing)
    EncoderIncoherent : BOOL;        // --> [SAFE] Incoherence ou hors bornes (FB_Encoder_Safety)
END_VAR
VAR_OUTPUT
    // === GATES DE FIABILITE ===
    EncoderFault      : BOOL;        // <-- [SAFE] Gate general fiabilite (SANS Homed) — vitesse/mouvements
    HomedAndReliable  : BOOL;        // <-- [STAT] Gate strict M3 : disponible ET reference ET pas incoherent
END_VAR

// 🛡️ 1. GATE GENERAL (D-A11, C1) — PAS de Homed : non-reference ≠ incoherent.
//    Ce gate sert a la fiabilite de la mesure (vitesse, mouvements, PositionsValid).
EncoderFault := (NOT EncoderAvailable) OR EncoderIncoherent;

// 🎯 2. GATE STRICT — reserve a l'interlock hauteur M3 (C1) : on ne translate pas
//    si la hauteur est inconnue (jamais home) ou douteuse.
HomedAndReliable := EncoderAvailable AND Homed AND (NOT EncoderIncoherent);
